(* IEC 61131-3 sources: SRCI_CLIENT_PLC/RobotLibrary/Library/Structures/Data, 1 file *)

(* ---- CyclicStateData.st ---- *)
{attribute 'pack_mode' := '1'}
// -------------------------------------------------------------------------
//  SRCI Robot Library
// -------------------------------------------------------------------------
//
//  Object:      CyclicStateData
//  Author:      Thorsten Brach
//  Date:        2024-06-01
//
//  Description:
//
//
//  Copyright:
//    (C) 2024 Thorsten Brach. All rights reserved
//             Licensed under the MIT License.
//
//  Disclaimer:
//    This project is provided without any guarantee and can be used for
//    private and commercial purposes. Any use is at the user’s
//    own risk and responsibility.
//
// -------------------------------------------------------------------------
TYPE CyclicStateData :
STRUCT
  /// Combination of various RA related states.
  StatusWord : RaStatusWord;
  /// Actual override in percentage multiplied by 100 (see chapter 5.6.2 for more information about the percentage encoding)
  Override   : UINT;
END_STRUCT
END_TYPE
